(* PLC project edge_two_sinks, ESBMC probe 1.0 *)
(* stored: creationDateTime 2026-10-07T00:00:00 *)

PROGRAM edge_two_sinks
  VAR_INPUT
    go : BOOL;
  END_VAR
  VAR_OUTPUT
    v : BOOL;
    b : BOOL;
  END_VAR
  VAR  (* added by the conversion: wires and edge detectors of the diagram *)
    R_TRIG1 : R_TRIG;
  END_VAR

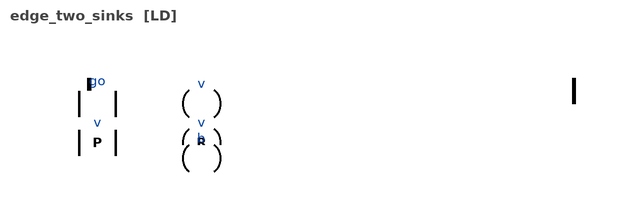
(* LD diagram, written out as Structured Text *)
v := go;
R_TRIG1(CLK := v);
IF R_TRIG1.Q THEN v := FALSE; END_IF;
b := R_TRIG1.Q;
END_PROGRAM

CONFIGURATION Config0
  RESOURCE Res0 ON PLC
    TASK tcyclic(INTERVAL := T#10ms, PRIORITY := 0);
    PROGRAM inst0 WITH tcyclic : edge_two_sinks;
  END_RESOURCE
END_CONFIGURATION
